Fanuc KAREL source: kb00109.KL

PROGRAM KB00109
%STACKSIZE=65535
%PRIORITY=65535
%NOLOCKGROUP
VAR
P1 : POSITION
RESULT : POSITION
BEGIN
-- UNRESOLVED_PC line 7 opcodes [27 22 1C 76 7E 4A] marker_code=0
END KB00109
